// TIA Portal V20 export
// export: Created 2026-10-19T18:06:33.9316453Z, ExportSetting WithDefaults, DisplayName Totally Integrated Automation Portal, DisplayVersion V20 Update 6, DisplayName TIA Portal Openness, DisplayVersion V20 Update 6, DisplayName TIA Portal Version Control Interface, DisplayVersion V20 Update 6, DisplayName SINAMICS Startdrive Advanced, DisplayVersion V20 SP1, DisplayName SINAMICS Startdrive G130, G150, S120, S150, SINAMICS MV, G220, S200, S210, DisplayVersion V20 SP1, DisplayName SINAMICS Startdrive G110M, G120, G120C, G120D, G120P, G115D, DisplayVersion V20 SP1, DisplayName STEP 7 Professional, DisplayVersion V20 Update 6, DisplayName STEP 7 Safety, DisplayVersion V20 Update 2, DisplayName WinCC Basic/Comfort/Advanced, DisplayVersion V20 Update 6, DisplayName WinCC Unified, DisplayVersion V20 Update 6
FUNCTION_BLOCK "SAI_IND_ZeroAdjust"   // FB52, LAD
TITLE = Zero Adjustment
{ S7_Optimized_Access := 'FALSE' }
VERSION : 0.1
// stored: AutoNumber true, IsIECCheckEnabled false, SetENOAutomatically false, UDAEnableTagReadback false
   VAR_INPUT
      ID : HW_IO;   // The Profinet Device Hardware Identifier under device properties
   END_VAR
   VAR_OUTPUT
      Process : Bool;   // Adjustment is in process
      Done : Bool;   // Adjustment completed successfully
      Error : Bool;
   END_VAR
   VAR_IN_OUT
      Start : Bool;   // Switch ON to start adjustment
   END_VAR
   VAR DB_SPECIFIC
      Activate : Bool;
      Status_RECORD : Int;
      Zero_RECORD : Int;
   END_VAR
   VAR
      WRREC_Zero { S7_SetPoint := 'True'} : WRREC;
      RDREC_Status { S7_SetPoint := 'True'} : RDREC;
   END_VAR
   VAR DB_SPECIFIC
      AdjustStep : SInt;
      Static01 : Bool;
      Static02 : Bool;
      Static03 : Bool;
   END_VAR
   VAR_TEMP   // added for the SCL form of the ladder/FBD networks
      _w1 : Bool;
      _w2 : Bool;
      _w3 : Bool;
      _w4 : Bool;
   END_VAR
BEGIN

REGION Network 1: Initialization
   // Initializes DONE and ERROR bits
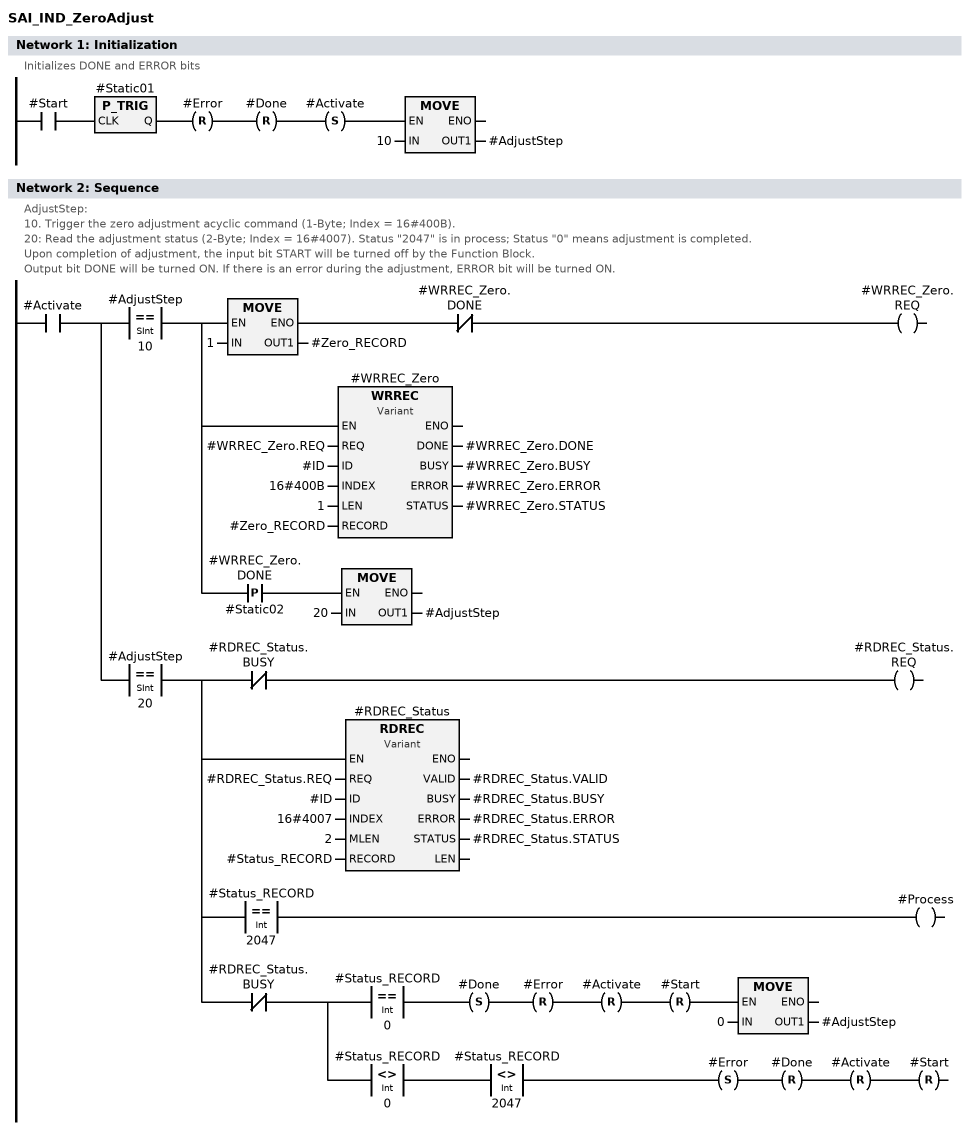
   RUNG wire#powerrail
      Contact( #Start )
      P_Trig( #Static01 )
      R_Coil( #Error )
      R_Coil( #Done )
      S_Coil( #Activate )
      { S7_GenerateENO := "TRUE" } Move(in := 10, out1 => #AdjustStep)
   END_RUNG
   // the same network as SCL:
   #_w1 := #Start AND NOT #Static01;   // rising edge
   #Static01 := #Start;
   IF #_w1 THEN
       #Error := FALSE;
       #Done := FALSE;
       #Activate := TRUE;
       #AdjustStep := 10;
   END_IF;
END_REGION

REGION Network 2: Sequence
   // AdjustStep:
   // 
   // 10. Trigger the zero adjustment acyclic command (1-Byte; Index = 16#400B). 
   // 
   // 20: Read the adjustment status (2-Byte; Index = 16#4007). Status "2047" is in process; Status "0" means adjustment is completed.
   // Upon completion of adjustment, the input bit START will be turned off by the Function Block.
   // Output bit DONE will be turned ON. If there is an error during the adjustment, ERROR bit will be turned ON.
   RUNG wire#powerrail
      Contact( #Activate )
      wire#w1
      { S7_Templates := "SrcType := SInt" } EQ_Contact(in1 := #AdjustStep, in2 := 10)
      wire#w2
      Move(in := 1, out1 => #Zero_RECORD)
      I_Contact( #WRREC_Zero.DONE )
      Coil( #WRREC_Zero.REQ )
   END_RUNG
   RUNG wire#w2
      { S7_Templates := "[ptr_type := Variant, id_type := HW_IO, index_type := DInt, len_type := UInt]" } #WRREC_Zero.WRREC(REQ := #WRREC_Zero.REQ, ID := #ID, INDEX := 16#400B, LEN := 1, RECORD := #Zero_RECORD, DONE => #WRREC_Zero.DONE, BUSY => #WRREC_Zero.BUSY, ERROR => #WRREC_Zero.ERROR, STATUS => #WRREC_Zero.STATUS)
   END_RUNG
   RUNG wire#w2
      P_Contact(operand := #WRREC_Zero.DONE, bit := #Static02)
      Move(in := 20, out1 => #AdjustStep)
   END_RUNG
   RUNG wire#w1
      { S7_Templates := "SrcType := SInt" } EQ_Contact(in1 := #AdjustStep, in2 := 20)
      wire#w3
      I_Contact( #RDREC_Status.BUSY )
      Coil( #RDREC_Status.REQ )
   END_RUNG
   RUNG wire#w3
      { S7_Templates := "[ptr_type := Variant, id_type := HW_IO, index_type := DInt, len_type := UInt]" } #RDREC_Status.RDREC(REQ := #RDREC_Status.REQ, ID := #ID, INDEX := 16#4007, MLEN := 2, RECORD := #Status_RECORD, VALID => #RDREC_Status.VALID, BUSY => #RDREC_Status.BUSY, ERROR => #RDREC_Status.ERROR, STATUS => #RDREC_Status.STATUS, LEN =>)
   END_RUNG
   RUNG wire#w3
      { S7_Templates := "SrcType := Int" } EQ_Contact(in1 := #Status_RECORD, in2 := 2047)
      Coil( #Process )
   END_RUNG
   RUNG wire#w3
      I_Contact( #RDREC_Status.BUSY )
      wire#w4
      { S7_Templates := "SrcType := Int" } EQ_Contact(in1 := #Status_RECORD, in2 := 0)
      S_Coil( #Done )
      R_Coil( #Error )
      R_Coil( #Activate )
      R_Coil( #Start )
      Move(in := 0, out1 => #AdjustStep)
   END_RUNG
   RUNG wire#w4
      { S7_Templates := "SrcType := Int" } NE_Contact(in1 := #Status_RECORD, in2 := 0)
      { S7_Templates := "SrcType := Int" } NE_Contact(in1 := #Status_RECORD, in2 := 2047)
      S_Coil( #Error )
      R_Coil( #Done )
      R_Coil( #Activate )
      R_Coil( #Start )
   END_RUNG
   // the same network as SCL:
   #_w1 := #Activate AND (#AdjustStep = 10);
   IF #_w1 THEN #Zero_RECORD := 1; END_IF;
   #WRREC_Zero.REQ := #_w1 AND NOT #WRREC_Zero.DONE;
   IF #_w1 THEN
       #WRREC_Zero(REQ := #WRREC_Zero.REQ,   // WRREC
                   ID := #ID,
                   INDEX := 16#400B,
                   LEN := 1,
                   RECORD := #Zero_RECORD,
                   DONE => #WRREC_Zero.DONE,
                   BUSY => #WRREC_Zero.BUSY,
                   ERROR => #WRREC_Zero.ERROR,
                   STATUS => #WRREC_Zero.STATUS);
   END_IF;
   #_w2 := #_w1 AND #WRREC_Zero.DONE AND NOT #Static02;   // rising edge of #WRREC_Zero.DONE
   #Static02 := #WRREC_Zero.DONE;
   IF #_w2 THEN #AdjustStep := 20; END_IF;
   #_w3 := #Activate AND (#AdjustStep = 20);
   #RDREC_Status.REQ := #_w3 AND NOT #RDREC_Status.BUSY;
   IF #_w3 THEN
       #RDREC_Status(REQ := #RDREC_Status.REQ,   // RDREC
                     ID := #ID,
                     INDEX := 16#4007,
                     MLEN := 2,
                     RECORD := #Status_RECORD,
                     VALID => #RDREC_Status.VALID,
                     BUSY => #RDREC_Status.BUSY,
                     ERROR => #RDREC_Status.ERROR,
                     STATUS => #RDREC_Status.STATUS);
   END_IF;
   #Process := #_w3 AND (#Status_RECORD = 2047);
   #_w4 := #_w3 AND NOT #RDREC_Status.BUSY;
   IF #_w4 AND (#Status_RECORD = 0) THEN
       #Done := TRUE;
       #Error := FALSE;
       #Activate := FALSE;
       #Start := FALSE;
       #AdjustStep := 0;
   END_IF;
   IF #_w4 AND (#Status_RECORD <> 0) AND (#Status_RECORD <> 2047) THEN
       #Error := TRUE;
       #Done := FALSE;
       #Activate := FALSE;
       #Start := FALSE;
   END_IF;
END_REGION
END_FUNCTION_BLOCK
